// SIMATIC S7-200 project (STEP 7-Micro/WIN), CPU 224 CN REL 02.01

SYMBOL_TABLE USUARIO1
SM2              I0.0     // Sensor magnetico extendido del cilindro retenedor
SM1              I0.1     // Sensor magnetico retraido del cilindor retenedor
SM4              I0.2     // Sensor magnetico extendido del cilindro de empuje
SM3              I0.3     // Sensor magnetico retraido del cilindor de empuje
SF               I0.4     // Sensor Fotoelectrico Final
SP               I0.5     // Sensor Fotoelectrico Superior
SP1              I0.6     // Sensor Fotoelectrico Inferior
SII              I0.7     // Sensor Inductivo
SB_1             I1.2     // Pulsador de marcha
SB_2             I1.3     // Pulsador de paro
QS               I1.4     // Zeta de Emergencia
SA               I1.5     // Selector de modo
KV1              Q0.0     // Cilindro neumatico Retenedor
KV2              Q0.1     // Cilindro neumatico de empuje
HL1              Q0.7     // Señalizacion amarillo
HL2              Q1.0     // Señalizacion verde
HL3              Q1.1     // Señalizacion roja
E0               M0.0     // Estado 0
E1               M0.1     // Estado 1
E2               M0.2     // Estado 2
E3               M0.3     // Estado 3
E4               M0.4     // Estado 4
E5               M0.5     // Estado 5
EM               M0.6     // Estado de emergencia
EP               M0.7     // Estado de parada
IN_UA            V3.0     // Bit de inicio
END_UA           V0.0     // Bit de finalizacion
SB1_UA           V3.1     // Pulsador de marcha
SB2_UA           V3.2     // Pulsador de parada
QS_UA            V3.3     // Zeta de emergencia
END_SYMBOL_TABLE

ORGANIZATION_BLOCK PRINCIPAL:OB1
TITLE=COMENTARIOS DEL PROGRAMA
BEGIN
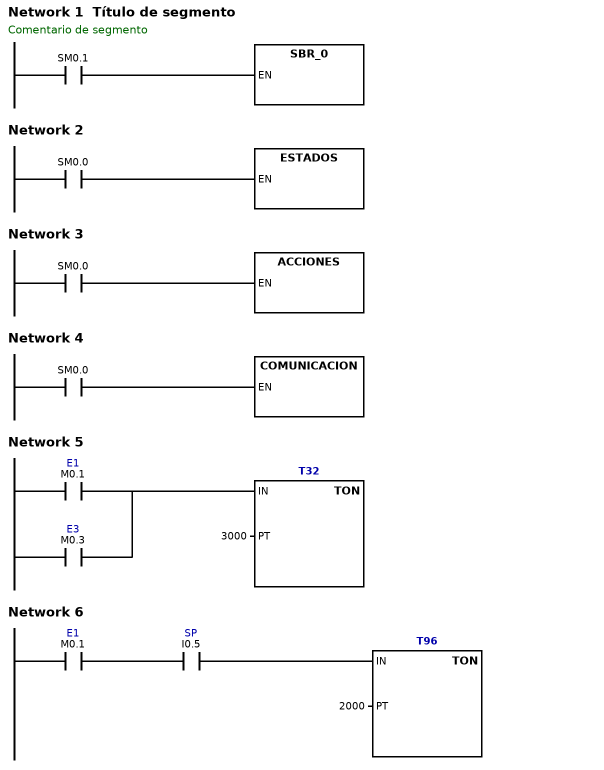
Network 1 // Título de segmento
// Comentario de segmento
LD     SM0.1
CALL   SBR_0:SBR0
Network 2
LD     SM0.0
CALL   ESTADOS:SBR1
Network 3
LD     SM0.0
CALL   ACCIONES:SBR2
Network 4
LD     SM0.0
CALL   COMUNICACION:SBR3
Network 5
LD     E1:M0.1
O      E3:M0.3
TON    T32, 3000
Network 6
LD     E1:M0.1
A      SP:I0.5
TON    T96, 2000
END_ORGANIZATION_BLOCK

SUBROUTINE_BLOCK SBR_0:SBR0
TITLE=COMENTARIOS DE LA SUBRUTINA
BEGIN
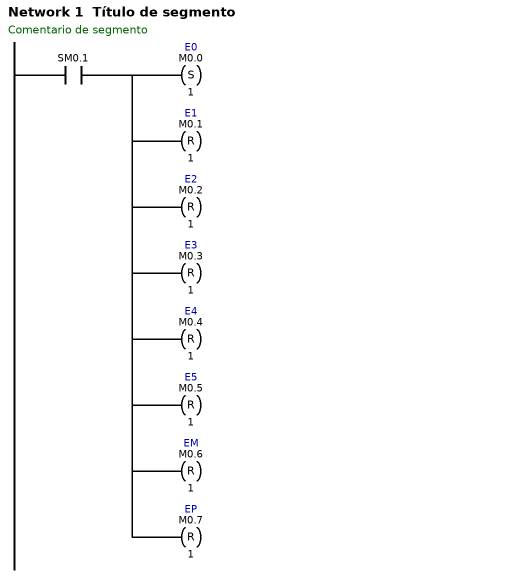
Network 1 // Título de segmento
// Comentario de segmento
LD     SM0.1
S      E0:M0.0, 1
R      E1:M0.1, 1
R      E2:M0.2, 1
R      E3:M0.3, 1
R      E4:M0.4, 1
R      E5:M0.5, 1
R      EM:M0.6, 1
R      EP:M0.7, 1
END_SUBROUTINE_BLOCK

SUBROUTINE_BLOCK ESTADOS:SBR1
TITLE=COMENTARIOS DE LA SUBRUTINA
BEGIN
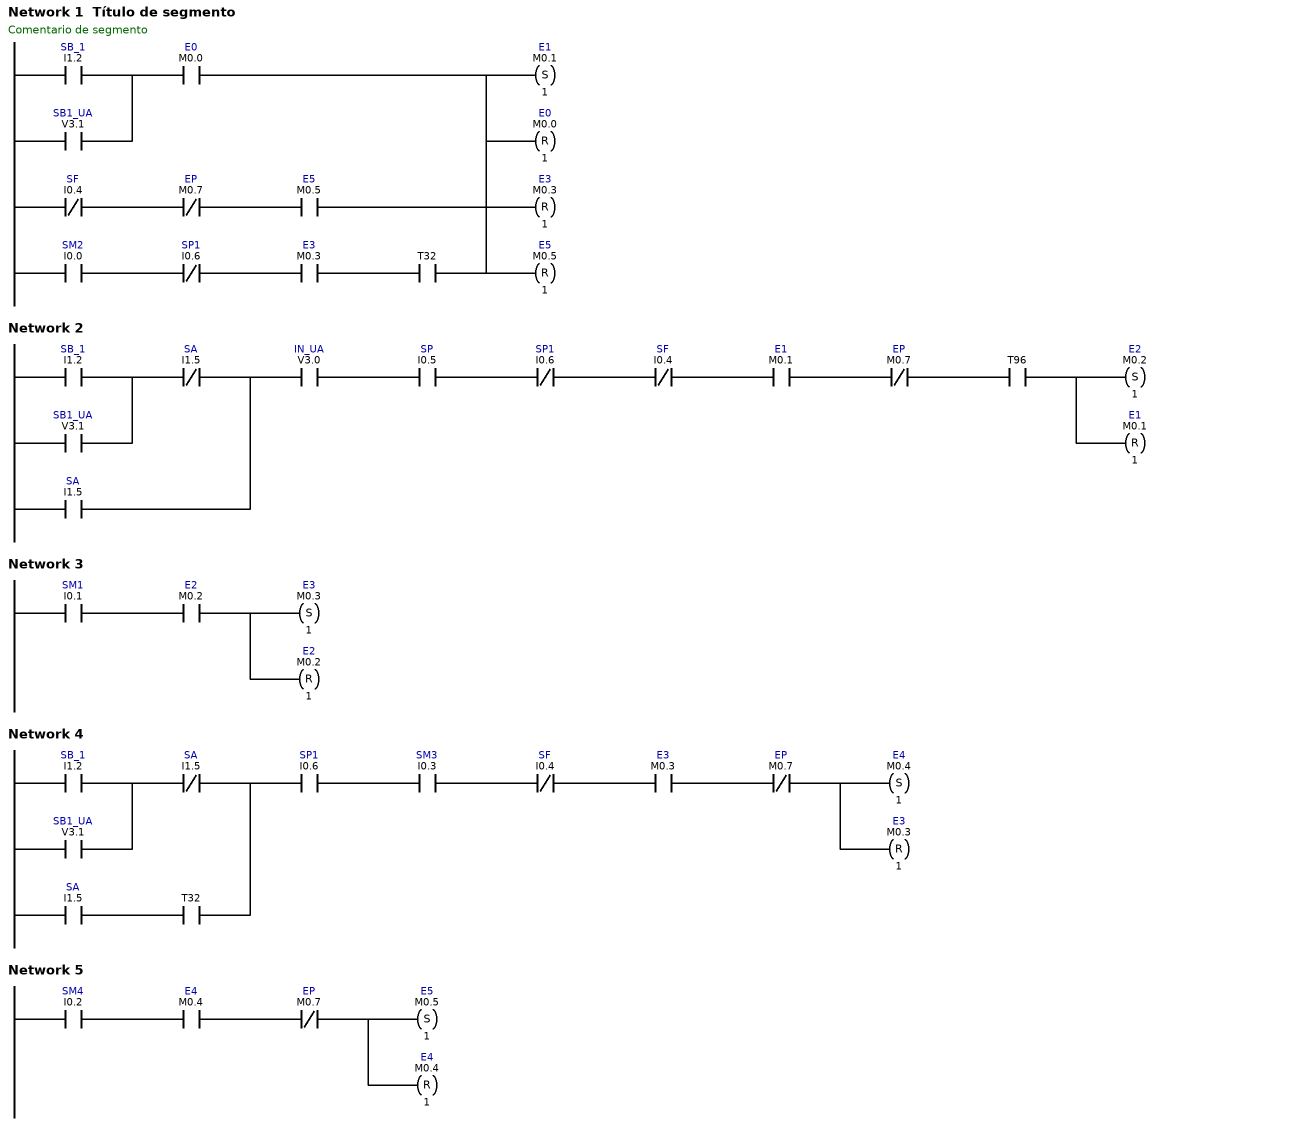
Network 1 // Título de segmento
// Comentario de segmento
LD     SB_1:I1.2
O      SB1_UA:V3.1
A      E0:M0.0
LDN    SF:I0.4
AN     EP:M0.7
A      E5:M0.5
LD     SM2:I0.0
AN     SP1:I0.6
A      E3:M0.3
A      T32
OLD
OLD
S      E1:M0.1, 1
R      E0:M0.0, 1
R      E3:M0.3, 1
R      E5:M0.5, 1
Network 2
LD     SB_1:I1.2
O      SB1_UA:V3.1
AN     SA:I1.5
O      SA:I1.5
A      IN_UA:V3.0
A      SP:I0.5
AN     SP1:I0.6
AN     SF:I0.4
A      E1:M0.1
AN     EP:M0.7
A      T96
S      E2:M0.2, 1
R      E1:M0.1, 1
Network 3
LD     SM1:I0.1
A      E2:M0.2
S      E3:M0.3, 1
R      E2:M0.2, 1
Network 4
LD     SB_1:I1.2
O      SB1_UA:V3.1
AN     SA:I1.5
LD     SA:I1.5
A      T32
OLD
A      SP1:I0.6
A      SM3:I0.3
AN     SF:I0.4
A      E3:M0.3
AN     EP:M0.7
S      E4:M0.4, 1
R      E3:M0.3, 1
Network 5
LD     SM4:I0.2
A      E4:M0.4
AN     EP:M0.7
S      E5:M0.5, 1
R      E4:M0.4, 1
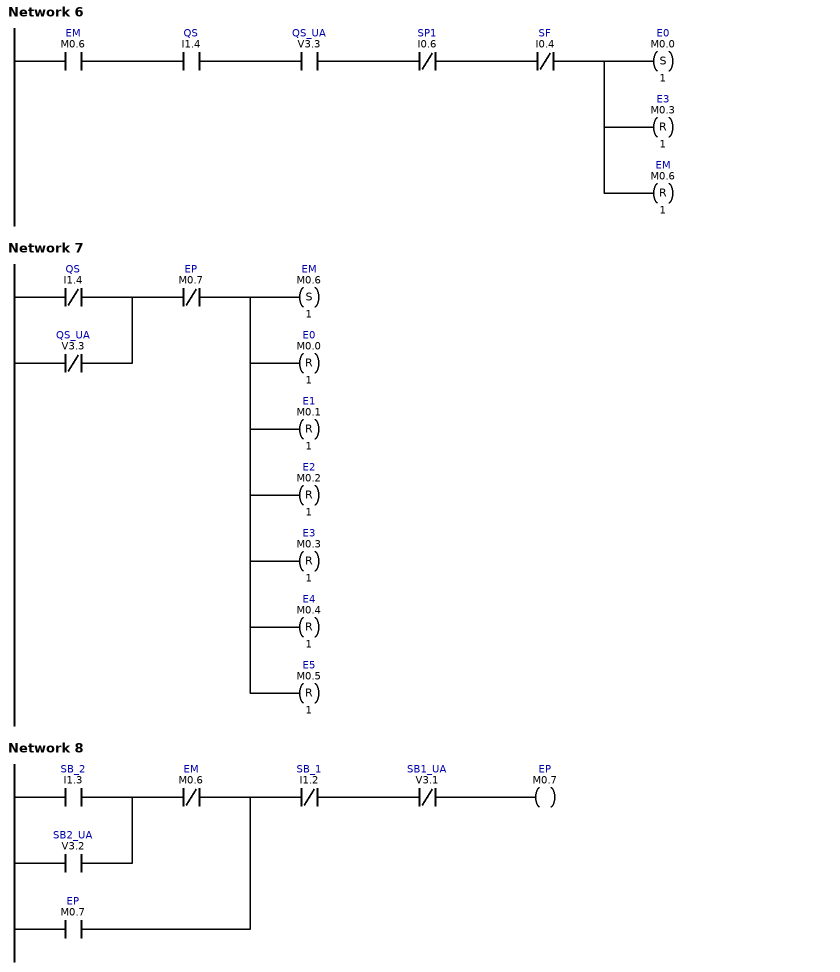
Network 6
// (network saved uncompiled; LAD cells follow)
// row 0: c0 -| |- EM:M0.6  c1 -| |- QS:I1.4  c2 -| |- QS_UA:V3.3  c3 -|/|- SP1:I0.6  c4 -|/|- SF:I0.4 v  c5 -(S) E0:M0.0, 1
// row 1: c4 ^v  c5 -(R) E3:M0.3, 1
// row 2: c4 ^  c5 -(R) EM:M0.6, 1
Network 7
LDN    QS:I1.4
ON     QS_UA:V3.3
AN     EP:M0.7
S      EM:M0.6, 1
R      E0:M0.0, 1
R      E1:M0.1, 1
R      E2:M0.2, 1
R      E3:M0.3, 1
R      E4:M0.4, 1
R      E5:M0.5, 1
Network 8
LD     SB_2:I1.3
O      SB2_UA:V3.2
AN     EM:M0.6
O      EP:M0.7
AN     SB_1:I1.2
AN     SB1_UA:V3.1
=      EP:M0.7
END_SUBROUTINE_BLOCK

SUBROUTINE_BLOCK ACCIONES:SBR2
TITLE=COMENTARIOS DE LA SUBRUTINA
BEGIN
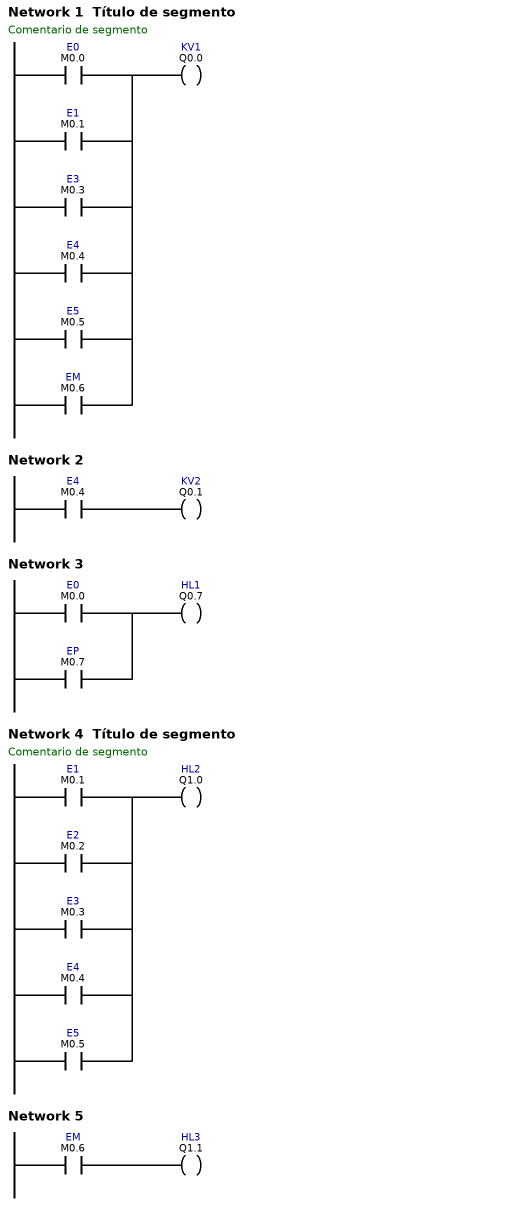
Network 1 // Título de segmento
// Comentario de segmento
LD     E0:M0.0
O      E1:M0.1
O      E3:M0.3
O      E4:M0.4
O      E5:M0.5
O      EM:M0.6
=      KV1:Q0.0
Network 2
LD     E4:M0.4
=      KV2:Q0.1
Network 3
LD     E0:M0.0
O      EP:M0.7
=      HL1:Q0.7
Network 4 // Título de segmento
// Comentario de segmento
LD     E1:M0.1
O      E2:M0.2
O      E3:M0.3
O      E4:M0.4
O      E5:M0.5
=      HL2:Q1.0
Network 5
LD     EM:M0.6
=      HL3:Q1.1
END_SUBROUTINE_BLOCK

SUBROUTINE_BLOCK COMUNICACION:SBR3
TITLE=COMENTARIOS DE LA SUBRUTINA
BEGIN
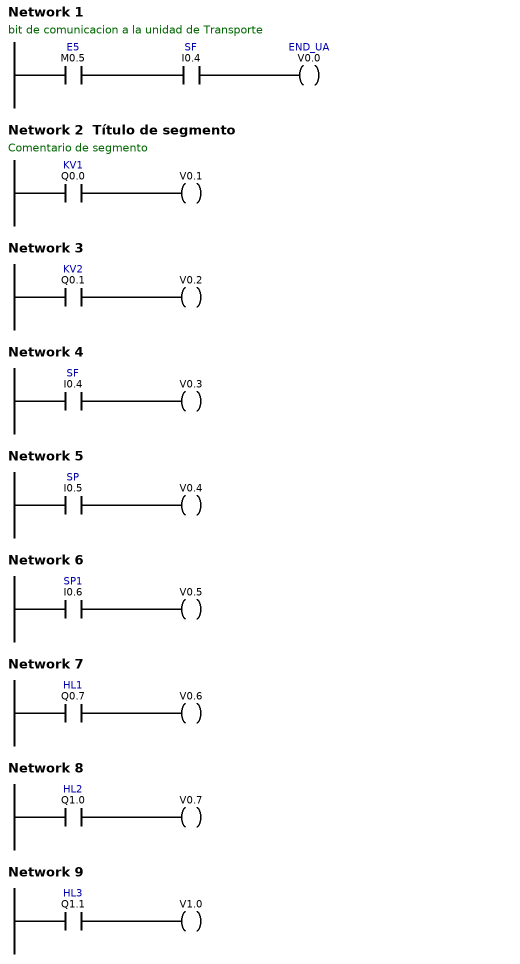
Network 1
// bit de comunicacion a la unidad de Transporte
LD     E5:M0.5
A      SF:I0.4
=      END_UA:V0.0
Network 2 // Título de segmento
// Comentario de segmento
LD     KV1:Q0.0
=      V0.1
Network 3
LD     KV2:Q0.1
=      V0.2
Network 4
LD     SF:I0.4
=      V0.3
Network 5
LD     SP:I0.5
=      V0.4
Network 6
LD     SP1:I0.6
=      V0.5
Network 7
LD     HL1:Q0.7
=      V0.6
Network 8
LD     HL2:Q1.0
=      V0.7
Network 9
LD     HL3:Q1.1
=      V1.0
END_SUBROUTINE_BLOCK
